(* IEC 61131-3 sources: plcassist-cli/packages/volt-lsp-iec/test-corpus/awa-palletizer/Device/Plc Logic/Application/Library Manager/CAA RTCLK, 8 files *)

(* ---- PROPERTYCONSTANTS.gvl ---- *)
VAR_GLOBAL
	GC_WTIMEZONESUPPORT : WORD := 1;
END_VAR

(* ---- VERSIONCONSTANTS.gvl ---- *)
VAR_GLOBAL
	GC_BYVERSION : BYTE := 1;
	GC_BYVERSION_1 : BYTE := 0;
END_VAR

(* ---- GETPROPERTY.fun ---- *)
FUNCTION GETPROPERTY : __XWORD
VAR_INPUT
	WPROPERTY : WORD;
END_VAR
END_FUNCTION

(* ---- GETSUPPLIERVERSION.fun ---- *)
FUNCTION GETSUPPLIERVERSION : WORD
VAR_INPUT
	XDUMMY : BOOL;
END_VAR
END_FUNCTION

(* ---- GETDATEANDTIME.fb ---- *)
FUNCTION_BLOCK GETDATEANDTIME
VAR_INPUT
	XEXECUTE : BOOL;
END_VAR
VAR_OUTPUT
	XDONE : BOOL;
	XBUSY : BOOL;
	XERROR : BOOL;
	EERROR : ERROR;
	DTDATEANDTIME : DATE_AND_TIME;
	ETIMEZONE : PERIODE;
END_VAR
VAR
	XPREVIOUSEXECUTE : BOOL;
	XPREVIOUSABORTINPROGRESS : BOOL;
	XABORTINPROGRESS : BOOL;
	IERROR : INT;
	HJOB : CAA.HANDLE;
	PGETDATEANDTIMEPARAMS : POINTER TO RTCLK_GETDATEANDTIME_PARAMS;
	STATEJOB : ASM.STATE;
	DWETRIGCLASS : __XWORD;
END_VAR
END_FUNCTION_BLOCK

METHOD FB_EXIT : BOOL
VAR_INPUT
	BINCOPYCODE : BOOL;
END_VAR
END_METHOD

METHOD FB_INIT : BOOL
VAR_INPUT
	BINITRETAINS : BOOL;
	BINCOPYCODE : BOOL;
END_VAR
END_METHOD

(* ---- GETTIMEZONEINFORMATION.fb ---- *)
FUNCTION_BLOCK GETTIMEZONEINFORMATION
VAR_INPUT
	XEXECUTE : BOOL;
END_VAR
VAR_OUTPUT
	XDONE : BOOL;
	XBUSY : BOOL;
	XERROR : BOOL;
	EERROR : ERROR;
	TZIINFO : RTCLK_TIME_ZONE_INFO;
END_VAR
VAR
	XPREVIOUSEXECUTE : BOOL;
	XPREVIOUSABORTINPROGRESS : BOOL;
	XABORTINPROGRESS : BOOL;
	IERROR : INT;
	HJOB : CAA.HANDLE;
	PGETTIMEZONEINFORMATIONPARAMS : POINTER TO RTCLK_GETTIMEZONEINFORMATION_PARAMS;
	STATEJOB : ASM.STATE;
	DWETRIGCLASS : __XWORD;
END_VAR
END_FUNCTION_BLOCK

METHOD FB_EXIT : BOOL
VAR_INPUT
	BINCOPYCODE : BOOL;
END_VAR
END_METHOD

METHOD FB_INIT : BOOL
VAR_INPUT
	BINITRETAINS : BOOL;
	BINCOPYCODE : BOOL;
END_VAR
END_METHOD

(* ---- SETDATEANDTIME.fb ---- *)
FUNCTION_BLOCK SETDATEANDTIME
VAR_INPUT
	XEXECUTE : BOOL;
	DTDATEANDTIME : DATE_AND_TIME;
END_VAR
VAR_OUTPUT
	XDONE : BOOL;
	XBUSY : BOOL;
	XERROR : BOOL;
	EERROR : ERROR;
END_VAR
VAR
	XPREVIOUSEXECUTE : BOOL;
	XPREVIOUSABORTINPROGRESS : BOOL;
	XABORTINPROGRESS : BOOL;
	IERROR : INT;
	HJOB : CAA.HANDLE;
	PSETDATEANDTIMEPARAMS : POINTER TO RTCLK_SETDATEANDTIME_PARAMS;
	STATEJOB : ASM.STATE;
	DWETRIGCLASS : __XWORD;
END_VAR
END_FUNCTION_BLOCK

METHOD FB_EXIT : BOOL
VAR_INPUT
	BINCOPYCODE : BOOL;
END_VAR
END_METHOD

METHOD FB_INIT : BOOL
VAR_INPUT
	BINITRETAINS : BOOL;
	BINCOPYCODE : BOOL;
END_VAR
END_METHOD

(* ---- SETTIMEZONEINFORMATION.fb ---- *)
FUNCTION_BLOCK SETTIMEZONEINFORMATION
VAR_INPUT
	XEXECUTE : BOOL;
	TZIINFO : RTCLK_TIME_ZONE_INFO;
END_VAR
VAR_OUTPUT
	XDONE : BOOL;
	XBUSY : BOOL;
	XERROR : BOOL;
	EERROR : ERROR;
END_VAR
VAR
	XPREVIOUSEXECUTE : BOOL;
	XPREVIOUSABORTINPROGRESS : BOOL;
	XABORTINPROGRESS : BOOL;
	IERROR : INT;
	HJOB : CAA.HANDLE;
	PSETTIMEZONEINFORMATIONPARAMS : POINTER TO RTCLK_SETTIMEZONEINFORMATION_PARAMS;
	STATEJOB : ASM.STATE;
	DWETRIGCLASS : __XWORD;
END_VAR
END_FUNCTION_BLOCK

METHOD FB_EXIT : BOOL
VAR_INPUT
	BINCOPYCODE : BOOL;
END_VAR
END_METHOD

METHOD FB_INIT : BOOL
VAR_INPUT
	BINITRETAINS : BOOL;
	BINCOPYCODE : BOOL;
END_VAR
END_METHOD
